(*
SPDX-FileCopyrightText: © 2026 Oleksandr Tiutyk <trofimich@gmail.com>
SPDX-License-Identifier: MIT
License: https://opensource.org/license/mit
*)

(*!
<summary>Runs the OpenFramework test groups registered by the shared test controller.</summary>
<description>
Owns persistent root instances and fixed child storage. The IO model group borrows the controller-owned fixture.
Use from one task without reentry.
Children borrows the same array for the instance lifetime. Root parents remain zero.
</description>
*)

{attribute 'no_assign'}
{attribute 'no_explicit_call' := 'do not call this function block directly'}
FUNCTION_BLOCK JsonConfigurationTestRunner EXTENDS TOF_Testing.TestRunner<45>
VAR_STAT
	//! <summary>Class name shared by instances of this concrete runner.</summary>
	{attribute 'hide'}
	_ClassName : STRING := __POUNAME();
END_VAR
VAR
	{attribute 'hide'}
	{attribute 'init_namespace'}
	_NamespaceName : STRING;
	//! <summary>Stable interface storage borrowed by the IO model group.</summary>
	_IOModelsFixture : IIOModelsTestFixture;
END_VAR
VAR_OUTPUT
	//! <summary>Owned root test suite for writer operations.</summary>
	WriterTest : JsonConfigurationWriterTest(name := "JsonConfigurationWriterTest", parent := 0);
	//! <summary>Owned root test suite for reader operations.</summary>
	ReaderTest : JsonConfigurationReaderTest(name := "JsonConfigurationReaderTest", parent := 0);
	//! <summary>Owned root test suite for round-trip serialization.</summary>
	RoundTripTest : JsonConfigurationRoundTripTest(name := "JsonConfigurationRoundTripTest", parent := 0);
	//! <summary>Owned root group for analog range conversions.</summary>
	RangeConverterTest : RangeAnalogValueConverterTest(name := "RangeAnalogValueConverterTest", parent := 0);
	//! <summary>Checks the two-cycle restart of an active timer.</summary>
	TimerRestartTest : TimerRestartWhileRunningTest(name := "RestartWhileRunning", parent := 0);
	//! <summary>Exercises failure to open a missing file for reading in an owned directory.</summary>
	MissingFileTest : OpenMissingFileForReadingTest(name := "OpenMissingFileForReading", parent := 0);
	//! <summary>Checks lexical file and directory path rules without filesystem I/O.</summary>
	PathValidationTest : LexicalPathValidationTest(name := "LexicalPathValidation", parent := 0);
	//! <summary>Groups the six filesystem contract tests that exercise no native I/O.</summary>
	FileSystemTests : FileSystemContractTest(name := "FileSystemContractTest", parent := 0);
	//! <summary>Groups the three native directory lifecycle scenarios.</summary>
	DirectoryTests : DirectoryTest(name := "DirectoryTest", parent := 0);
	//! <summary>Groups the four cyclic file-content manager scenarios.</summary>
	FileContentTests : FileContentManagerOperationsTest(name := "FileContentManagerTest", parent := 0);
	//! <summary>Groups the three native filesystem integration scenarios.</summary>
	FileSystemIntegrationTests : FileSystemIntegrationTestGroup(name := "FileSystemIntegrationTest", parent := 0);
	//! <summary>Groups the deterministic logger contracts and task-routing tests.</summary>
	LoggerContractTests : LoggerContractTestGroup(name := "LoggerContractTest", parent := 0);
	//! <summary>Runs the native file and EventLogger integration cases.</summary>
	LoggerIntegrationTests : LoggerIntegrationTestGroup(name := "LoggerTest", parent := 0);
	//! <summary>Groups the task lifecycle view and naming cases.</summary>
	TaskLifecycleTests : TaskLifecycleViewsTestGroup(name := "TaskLifecycleViewsTest", parent := 0);
	//! <summary>Groups FIFO and empty-queue behavior.</summary>
	TaskSequenceTests : TaskSequenceTestGroup(name := "TaskSequenceTest", parent := 0);
	//! <summary>Groups cooperative queue cleanup and failure cases.</summary>
	TaskQueueCleanupTests : TaskQueueCleanupTestGroup(name := "TaskQueueCleanupTest", parent := 0);
	//! <summary>Groups timer timing, lifecycle and restart cases.</summary>
	TimerTimingTests : TimerTimingTestGroup(name := "TimerTimingTest", parent := 0);
	//! <summary>Groups task stopping, failure and naming cases.</summary>
	TaskStoppingTests : TaskStoppingTestGroup(name := "TaskStoppingTest", parent := 0);
	//! <summary>Groups concrete object disposal and address conversion cases.</summary>
	ObjectLifetimeTests : ObjectLifetimeTestGroup(name := "ObjectLifetimeTest", parent := 0);
	//! <summary>Groups generic storage, ordering, conversion and runtime type diagnostics.</summary>
	GenericValueTests : GenericValueTestGroup(name := "GenericValueTest", parent := 0);
	//! <summary>Groups random range and dispersion contracts.</summary>
	RandomTests : RandomTestGroup(name := "RandomTest", parent := 0);
	//! <summary>Groups exception transport, cloning, diagnostics and failure boundaries.</summary>
	ExceptionTests : ExceptionTestGroup(name := "ExceptionTest", parent := 0);
	//! <summary>Groups byte-string formatting, editing, search and splitter contracts.</summary>
	StringTests : StringsTestGroup(name := "StringsTest", parent := 0);
	//! <summary>Groups wide-string formatting, editing, search and splitter contracts.</summary>
	WideStringTests : WideStringsTestGroup(name := "WideStringsTest", parent := 0);
	//! <summary>Groups byte-string builder assignment, reuse and failure contracts.</summary>
	StringBuilderTests : StringBuilderTestGroup(name := "StringBuilderTest", parent := 0);
	//! <summary>Groups wide-string builder assignment, reuse and failure cases.</summary>
	WideStringBuilderTests : WideStringBuilderTestGroup(name := "WideStringBuilderTest", parent := 0);
	//! <summary>Groups byte-list operations with dynamically allocated storage.</summary>
	DynamicByteListTests : DynamicByteListTestGroup(name := "DynamicByteListTest", parent := 0);
	//! <summary>Groups fixed-capacity byte-list operations and overflow handling.</summary>
	StaticByteListTests : StaticByteListTestGroup(name := "StaticByteListTest", parent := 0);
	//! <summary>Groups native JSON conversion, capacity, encoding and callback cases.</summary>
	AutomaticJsonSerializerTests : AutomaticJsonSerializerTestGroup(name := "AutomaticJsonSerializerTest", parent := 0);
	//! <summary>Groups fixed-capacity queue lookup, FIFO, clear and overflow cases.</summary>
	StaticQueueTests : StaticQueueTestGroup(name := "StaticQueueTest", parent := 0);
	//! <summary>Groups dynamic queue lookup, FIFO, growth and clear cases.</summary>
	DynamicQueueTests : DynamicQueueTestGroup(name := "DynamicQueueTest", parent := 0);
	//! <summary>Groups dynamic dictionary lookup, update, removal and clear cases.</summary>
	DynamicDictionaryTests : DynamicDictionaryTestGroup(name := "DynamicDictionaryTest", parent := 0);
	//! <summary>Groups fixed-capacity dictionary lookup, update, removal, clear and overflow cases.</summary>
	StaticDictionaryTests : StaticDictionaryTestGroup(name := "StaticDictionaryTest", parent := 0);
	//! <summary>Groups dynamic set lookup, duplicate updates, removal and clear cases.</summary>
	DynamicUniqueDataSetTests : DynamicUniqueDataSetTestGroup(name := "DynamicUniqueDataSetTest", parent := 0);
	//! <summary>Groups fixed-capacity set lookup, duplicate updates, removal, clear and overflow cases.</summary>
	StaticUniqueDataSetTests : StaticUniqueDataSetTestGroup(name := "StaticUniqueDataSetTest", parent := 0);
	//! <summary>Groups dynamic list copying, borrowing, editing, search, sorting and clear cases.</summary>
	DynamicListTests : DynamicListTestGroup(name := "DynamicListTest", parent := 0);
	//! <summary>Groups fixed-capacity list copying, borrowing, editing, search, sorting and overflow cases.</summary>
	StaticListTests : StaticListTestGroup(name := "StaticListTest", parent := 0);
	//! <summary>Groups dynamic stack storage, LIFO order, cursors and ownership cases.</summary>
	DynamicStackTests : DynamicStackTestGroup(name := "DynamicStackTest", parent := 0);
	//! <summary>Groups fixed-capacity stack storage, LIFO order, cursors, ownership and overflow cases.</summary>
	StaticStackTests : StaticStackTestGroup(name := "StaticStackTest", parent := 0);
	//! <summary>Groups digital and analog device, simulated channel and conversion cases.</summary>
	DevicesIOTests : DevicesIOTestGroup(name := "DevicesIOTest", parent := 0);
	//! <summary>Groups collection ownership, callback, growth and enumeration scenarios.</summary>
	CollectionsContractTests : CollectionsContractTestGroup(name := "CollectionsContractTest", parent := 0);
	//! <summary>Groups PDO representation and simulated input binding scenarios.</summary>
	IOModelsTests : IOModelsTestGroup(name := "IOModelsTest", parent := 0, fixtureSlot := ADR(_IOModelsFixture));
	//! <summary>Groups workflow integration, comparison and variable-scope scenarios.</summary>
	WorkflowComprehensiveTests : WorkflowComprehensiveTestGroup(name := "WorkflowComprehensiveTest", parent := 0);
	//! <summary>Groups workflow contracts and the cyclic delay timing regression.</summary>
	WorkflowContractTests : WorkflowContractTestGroup(name := "WorkflowContractTest", parent := 0);
	//! <summary>Groups automation component contracts and observations from the dedicated runner task.</summary>
	AutomationComponentTests : AutomationComponentTestGroup(name := "AutomationComponentTest", parent := 0);
END_VAR
VAR
	_Children : ARRAY [0.._ChildCount - 1] OF TOF_Testing.ITestElement :=
	[
		WriterTest,
		ReaderTest,
		RoundTripTest,
		RangeConverterTest,
		TimerRestartTest,
		MissingFileTest,
		PathValidationTest,
		FileSystemTests,
		DirectoryTests,
		FileContentTests,
		FileSystemIntegrationTests,
		LoggerContractTests,
		LoggerIntegrationTests,
		TaskLifecycleTests,
		TaskSequenceTests,
		TaskQueueCleanupTests,
		TimerTimingTests,
		TaskStoppingTests,
		ObjectLifetimeTests,
		GenericValueTests,
		RandomTests,
		ExceptionTests,
		StringTests,
		WideStringTests,
		StringBuilderTests,
		WideStringBuilderTests,
		DynamicByteListTests,
		StaticByteListTests,
		AutomaticJsonSerializerTests,
		StaticQueueTests,
		DynamicQueueTests,
		DynamicDictionaryTests,
		StaticDictionaryTests,
		DynamicUniqueDataSetTests,
		StaticUniqueDataSetTests,
		DynamicListTests,
		StaticListTests,
		DynamicStackTests,
		StaticStackTests,
		DevicesIOTests,
		CollectionsContractTests,
		IOModelsTests,
		WorkflowComprehensiveTests,
		WorkflowContractTests,
		AutomationComponentTests
	];
END_VAR

(*!
<summary>Stores the controller-owned model fixture for the IO model group.</summary>
<description>Stores a borrow without invoking the fixture. The controller keeps it alive for all test runs.</description>
<param name="ioModelsFixture">Controller-owned model fixture declared before the runner.</param>
*)
METHOD FB_init : BOOL
VAR_INPUT
	bInitRetains: BOOL; // TRUE: the retain variables are initialized (reset warm / reset cold)
	bInCopyCode: BOOL; // TRUE: the instance will be copied to the copy code afterward (online change)
	ioModelsFixture : IIOModelsTestFixture;
END_VAR
IF NOT bInCopyCode THEN
	_IOModelsFixture := ioModelsFixture;
END_IF

FB_init := TRUE;
END_METHOD

(*!
<summary>Borrows the unchanged persistent root array; application code must not modify it.</summary>
*)
{attribute 'monitoring' := 'call'}
PROPERTY Children : REFERENCE TO ARRAY [0.._ChildCount - 1] OF TOF_Testing.ITestElement
GET
Children REF= _Children;
END_GET
END_PROPERTY

(*!
<summary>Borrows the concrete class name; callers must not modify the returned storage.</summary>
*)
{attribute 'monitoring' := 'call'}
PROPERTY ClassName : REFERENCE TO STRING
GET
ClassName REF= _ClassName;
END_GET
END_PROPERTY

(*!
<summary>Borrows the concrete namespace name for the instance lifetime; callers must not modify it.</summary>
*)
{attribute 'monitoring' := 'call'}
PROPERTY NamespaceName : REFERENCE TO STRING
GET
NamespaceName REF= _NamespaceName;
END_GET
END_PROPERTY

(*!
<summary>Reports the complete concrete instance size in bytes.</summary>
*)
{attribute 'monitoring' := 'call'}
PROPERTY SelfSize : ULINT
GET
SelfSize := XSIZEOF(THIS^);
END_GET
END_PROPERTY

END_FUNCTION_BLOCK

(* stored: Version 1.1.0.1
   POU JsonConfigurationTestRunner: Id {6cc84da6-ca7e-4045-bc76-1f4d20ac227c}, SpecialFunc None
   Method FB_init: Id {a83b8d0d-6f01-4243-a28c-ccae384cb4c1}
   Property Children: Id {31c7bfc8-0e68-4e3e-a176-58572bbcdaa1}
   Get Get: Id {512b21ae-1365-4e94-a4cc-90a7092ed49b}
   Property ClassName: Id {80c87378-a184-4f48-8fa4-8458bfb9bc53}
   Get Get: Id {37612fee-83d8-4ac2-aae0-486db11c1c15}
   Property NamespaceName: Id {944543d8-d3b3-4c53-b852-c12c99129d33}
   Get Get: Id {7340f8de-5251-4a6e-af92-3c555dabd6dc}
   Property SelfSize: Id {986cda70-ca4c-4ad3-bf14-98d5e09ecaf8}
   Get Get: Id {c07881e0-fcd6-46ff-826a-c9dd1bdfd319} *)
